{attribute 'qualified_only'}
VAR_GLOBAL
	Q1_Actual : LREAL;
    Q2_Actual : LREAL;
    Q3_Actual : LREAL;
END_VAR

(* stored: Version 1.1.0.1, ProductVersion 3.1.4024.15
   GVL GVL_RobotData: Id {0106388c-f998-44c0-a906-c16ba42ce6ae} *)
